TYPE "ST_CylinderDevice"
VERSION : 0.1
   STRUCT
      Direction : DInt;
      Withdrawn : Bool;
      Extended : Bool;
      Retracted : Bool;
      Lease : "ST_SequenceCommandLease";
   END_STRUCT;

END_TYPE

